(* IEC 61131-3 sources: ia2/examples/tier0-control/sim/pous, 1 file *)

(* ---- main.st ---- *)
PROGRAM main
VAR
    sp_flow : REAL;
    big : DINT;
    lamp : BOOL;
    ticks : UDINT := 0;
END_VAR
ticks := (ticks + 1) MOD 1000000000;
END_PROGRAM
